(* IEC 61131-3 sources: vscode-twincat-st/src/sample/Base/DUTs, 4 files *)

(* ---- Aliases.st ---- *)
TYPE MyAlias : USINT;
END_TYPE

(* ---- Enums.st ---- *)
TYPE MyEnum1 :
(
    White := 0
);
END_TYPE

TYPE MyEnum2 :
(
    White   := 0,

    Yellow  := 1
) DWORD := Yellow;
END_TYPE

TYPE INTERNAL MyEnum3 :
(
    White := 0,

    Yellow
) DWORD;
END_TYPE

TYPE MyEnum4 :
(
    White := 0
) := White;
END_TYPE

(* ---- Structs.st ---- *)
TYPE MyStruct :
STRUCT
    A: BOOL;

    B: INT;

	C: BOOL := 1;
END_STRUCT
END_TYPE

(* ---- Unions.st ---- *)
TYPE MyUnion:
UNION
    A: LREAL;

    B: LINT;

    C: WORD := 1;
END_UNION
END_TYPE
